(* IEC 61131-3 sources: tsplc/packages/vscode-extension/tests/fixtures/conveyor/types, 3 files *)

(* ---- ST_Conveyor.st ---- *)
TYPE ST_Conveyor :
STRUCT
	ZoneCount : UINT;
	Zones : ARRAY[1..128] OF ST_Zone;
END_STRUCT
END_TYPE

(* ---- ST_Output.st ---- *)
TYPE ST_Output :
STRUCT
	MotionAsserted : BOOL;
	Speed : UINT;
END_STRUCT
END_TYPE

(* ---- ST_Zone.st ---- *)
TYPE ST_Zone :
STRUCT
	Output : ST_Output;
	Ready : BOOL;
END_STRUCT
END_TYPE
